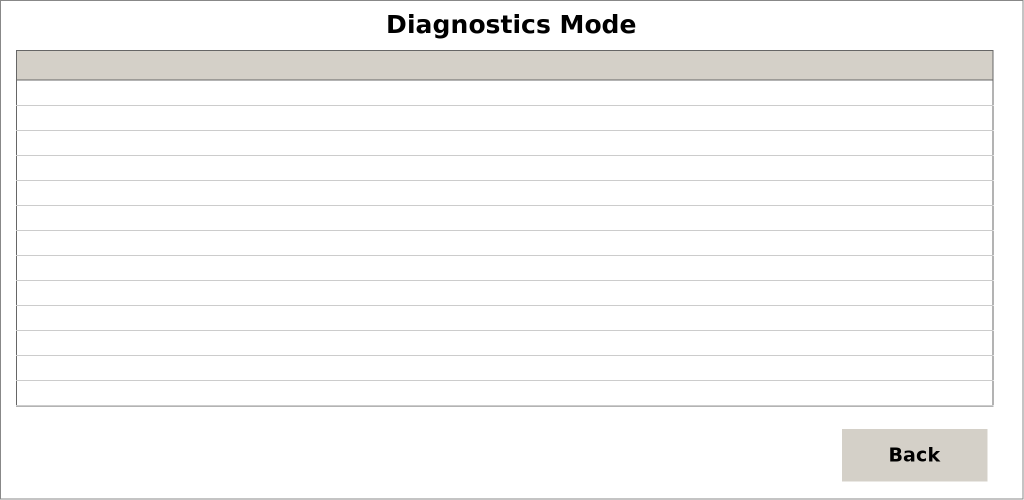
VISUALIZATION V_Diagnostics  // 1024x500
VAR_IN_OUT
Machine_HMI : ST_Machine_HMI;
END_VAR
    Label (0,-1 1023x50), "Diagnostics Mode"
    Table (16,50 977x356), data array: MAIN.Seedra.Machine_HMI.aAlarmHistory
        p338671338: MAIN.Seedra.Machine_HMI.aAlarmHistory[INDEX].sMessageText
        p1892666644: MAIN.Seedra.Machine_HMI.aAlarmHistory[INDEX].nTimestamp
        p3854506369: MAIN.Seedra.Machine_HMI.aAlarmHistory[INDEX].eSeverity
    RoundedRectangle (842,429 145x52), "Back"
        OnMouseUp: execute { GVL_HMI.PopupToDisplay := 0; }
END_VISUALIZATION

(* stored: Version 1.1.0.1, ProductVersion 3.1.4024.15
   Visu V_Diagnostics: Id {210d888d-4f35-4c7d-92f4-67383adc7a80} *)
